(* PLC project boton_matriz, UCuenca DEET Tablero DEET 1 *)
(* stored: creationDateTime 2026-10-19T12:00:00, modificationDateTime 2026-10-19T12:00:00 *)

(* Mientras pulsas I16 se encienden las 9 luces de la matriz 3x3. *)
PROGRAM boton_matriz
  VAR
    BOTON AT %IX102.0 : BOOL;  (* Pulsador I16 del Controllino *)
    D0 AT %QX100.0 : BOOL;  (* Luz D0 de la matriz *)
    D1 AT %QX100.1 : BOOL;  (* Luz D1 de la matriz *)
    D2 AT %QX100.2 : BOOL;  (* Luz D2 de la matriz *)
    D6 AT %QX100.6 : BOOL;  (* Luz D6 de la matriz *)
    D7 AT %QX100.7 : BOOL;  (* Luz D7 de la matriz *)
    D8 AT %QX101.0 : BOOL;  (* Luz D8 de la matriz *)
    D12 AT %QX101.4 : BOOL;  (* Luz D12 de la matriz *)
    D13 AT %QX101.5 : BOOL;  (* Luz D13 de la matriz *)
    D14 AT %QX101.6 : BOOL;  (* Luz D14 de la matriz *)
  END_VAR

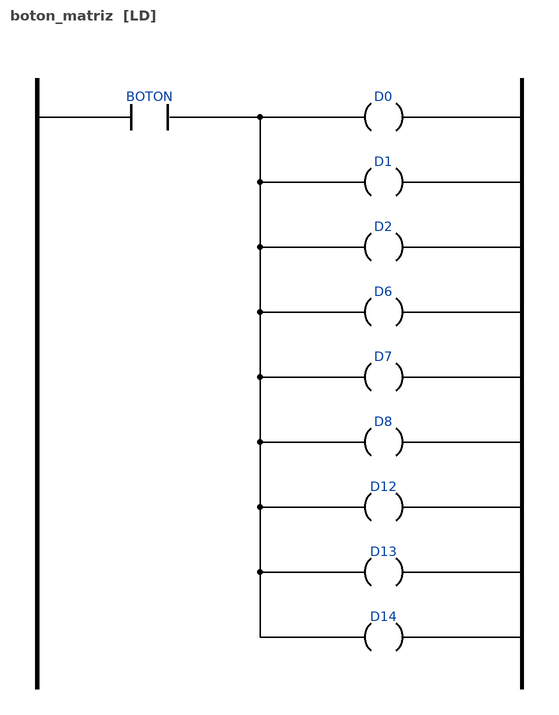
(* LD diagram, written out as Structured Text *)
D0 := BOTON;
D1 := BOTON;
D2 := BOTON;
D6 := BOTON;
D7 := BOTON;
D8 := BOTON;
D12 := BOTON;
D13 := BOTON;
D14 := BOTON;
END_PROGRAM

CONFIGURATION Config0
  RESOURCE Res0 ON PLC
    TASK task0(INTERVAL := T#20ms, PRIORITY := 0);
    PROGRAM instance0 WITH task0 : boton_matriz;
  END_RESOURCE
END_CONFIGURATION
